(* IEC 61131-3 sources: rusty/tests/lit/multi/external_unit_linkage, 25 files *)

(* ---- interfaces_main.st ---- *)
FUNCTION main : DINT
VAR
    fa : FbA;
    fb : FbB;
END_VAR
    printf('%d$N', call_a(fa));
    printf('%d$N', call_b(fb));
END_FUNCTION

(* ---- properties_c_main.st ---- *)
FUNCTION main : DINT
VAR
    fb : FbExt;
END_VAR
    fb.value := 42;
    printf('%d$N', fb.value);
    printf('%d$N', fb.getValue());
END_FUNCTION

(* ---- properties_main.st ---- *)
FUNCTION main : DINT
VAR
    base : FbBase;
    child : FbChild;
    counter : Counter;
    iface : IValue;
END_VAR
    base.value := 42;
    printf('%d$N', base.value);

    child.value := 5;
    printf('%d$N', child.value);

    printf('%d$N', counter.count);

    iface := child;
    printf('%d$N', iface.value);
END_FUNCTION

(* ---- reference_to_return_lib.st ---- *)
FUNCTION increment : REFERENCE TO DINT
VAR_INPUT
    value : REFERENCE TO DINT;
END_VAR
    value := value + 1;
    increment REF= value;
END_FUNCTION

FUNCTION increment_twice : DINT
VAR
    x : DINT := 5;
    r : REFERENCE TO DINT;
END_VAR
    r REF= x;
    r REF= increment(r);
    r REF= increment(r);
    increment_twice := r;
END_FUNCTION

(* ---- reference_to_return_main.st ---- *)
FUNCTION main : DINT
VAR
    x : DINT := 2;
    r : REFERENCE TO DINT;
END_VAR
    r REF= x;
    r REF= increment(r);
    printf('%d$N', r);
    printf('%d$N', increment_twice());
END_FUNCTION

(* ---- retain_main.st ---- *)
FUNCTION main : DINT
    RetainProgram();
    printf('%d$N', RetainProgram.count);
    printf('%d$N', retainFb.value);
END_FUNCTION

(* ---- retained_fat_pointer_main.st ---- *)
FUNCTION main
    bindA();
    bindB();
    consumerA();
    consumerB();
    printf('%d %d$N', consumerA.result, consumerB.result);
END_FUNCTION

(* ---- retained_fat_pointer_overload_main.st ---- *)
FUNCTION main
    // CHECK: main: done
    printf('main: done$N');
END_FUNCTION

(* ---- retained_fat_pointer_property_main.st ---- *)
FUNCTION main
    VAR
        ownerA : OwnerA;
        ownerB : OwnerB;
    END_VAR
    printf('%d %d$N', ownerA.value, ownerB.value);
END_FUNCTION

(* ---- interface_dispatch_lib.st ---- *)
INTERFACE IShape
    METHOD area : DINT END_METHOD
    PROPERTY_GET name : DINT END_PROPERTY
END_INTERFACE

INTERFACE ISolid EXTENDS IShape
    METHOD volume : DINT END_METHOD
END_INTERFACE

INTERFACE ILogger
    METHOD log : DINT
    VAR_INPUT value : DINT; END_VAR
    END_METHOD
END_INTERFACE

FUNCTION_BLOCK LibSquare IMPLEMENTS IShape
VAR
    side : DINT := 3;
END_VAR
    METHOD area : DINT area := side * side; END_METHOD
    PROPERTY_GET name : DINT name := 100; END_PROPERTY
END_FUNCTION_BLOCK

FUNCTION_BLOCK LibCube EXTENDS LibSquare IMPLEMENTS ISolid
    METHOD volume : DINT volume := area() * side; END_METHOD
    PROPERTY_GET name : DINT name := 200; END_PROPERTY
END_FUNCTION_BLOCK

FUNCTION lib_area_of : DINT
VAR_INPUT shape : IShape; END_VAR
    lib_area_of := shape.area() + shape.name;
END_FUNCTION

FUNCTION_BLOCK LibService
VAR
    logger : ILogger;
    shapes : ARRAY[0..1] OF IShape;
END_VAR
    METHOD inject
    VAR_INPUT l : ILogger; END_VAR
        logger := l;
    END_METHOD

    METHOD add_shape
    VAR_INPUT i : DINT; s : IShape; END_VAR
        shapes[i] := s;
    END_METHOD

    METHOD run : DINT
        run := logger.log(shapes[0].area() + shapes[1].area());
    END_METHOD
END_FUNCTION_BLOCK

FUNCTION lib_volume_as_shape : DINT
VAR_INPUT solid : ISolid; END_VAR
VAR shape : IShape; END_VAR
    shape := solid;
    lib_volume_as_shape := solid.volume() + shape.area();
END_FUNCTION

(* ---- interface_dispatch_main.st ---- *)
FUNCTION_BLOCK AppLogger IMPLEMENTS ILogger
VAR
    last : DINT;
END_VAR
    METHOD log : DINT
    VAR_INPUT value : DINT; END_VAR
        last := value;
        log := value + 1;
    END_METHOD
END_FUNCTION_BLOCK

FUNCTION_BLOCK AppCircle IMPLEMENTS IShape
    METHOD area : DINT area := 7; END_METHOD
    PROPERTY_GET name : DINT name := 300; END_PROPERTY
END_FUNCTION_BLOCK

FUNCTION_BLOCK AppBigCube EXTENDS LibCube
    METHOD area : DINT area := 50; END_METHOD
END_FUNCTION_BLOCK

FUNCTION main : DINT
VAR
    square : LibSquare;
    cube : LibCube;
    bigCube : AppBigCube;
    circle : AppCircle;
    logger : AppLogger;
    service : LibService;
    shape : IShape;
    solid : ISolid;
END_VAR
    // Lib type, called through an interface in the app
    shape := square;
    printf('%d %d$N', shape.area(), shape.name);
    shape := cube;
    printf('%d %d$N', shape.area(), shape.name);
    solid := cube;
    printf('%d$N', solid.volume());

    // App type passed to a lib function that calls through the interface
    printf('%d$N', lib_area_of(circle));
    printf('%d$N', lib_area_of(square));

    // App type that extends a lib type, overriding a method
    shape := bigCube;
    printf('%d %d$N', shape.area(), shape.name);
    printf('%d$N', lib_volume_as_shape(bigCube));

    // Dependency inversion: the lib stores app objects and calls them later
    service.inject(logger);
    service.add_shape(0, circle);
    service.add_shape(1, bigCube);
    printf('%d %d$N', service.run(), logger.last);
END_FUNCTION

(* ---- interfaces_lib_a.st ---- *)
INTERFACE IA
    METHOD a : DINT END_METHOD
END_INTERFACE

FUNCTION_BLOCK FbA IMPLEMENTS IA
    METHOD a : DINT
        a := 1;
    END_METHOD
END_FUNCTION_BLOCK

FUNCTION call_a : DINT
VAR_INPUT
    x : IA;
END_VAR
    call_a := x.a();
END_FUNCTION

(* ---- interfaces_lib_b.st ---- *)
INTERFACE IB
    METHOD b : DINT END_METHOD
END_INTERFACE

FUNCTION_BLOCK FbB IMPLEMENTS IB
    METHOD b : DINT
        b := 2;
    END_METHOD
END_FUNCTION_BLOCK

FUNCTION call_b : DINT
VAR_INPUT
    x : IB;
END_VAR
    call_b := x.b();
END_FUNCTION

(* ---- properties_lib.st ---- *)
INTERFACE IValue
    PROPERTY_GET value : DINT END_PROPERTY
END_INTERFACE

FUNCTION_BLOCK FbBase IMPLEMENTS IValue
VAR
    _value : DINT;
END_VAR
    PROPERTY_GET value : DINT
        value := _value;
    END_PROPERTY

    PROPERTY_SET value : DINT
        _value := value;
    END_PROPERTY
END_FUNCTION_BLOCK

FUNCTION_BLOCK FbChild EXTENDS FbBase
    PROPERTY_GET value : DINT
        value := _value * 2;
    END_PROPERTY
END_FUNCTION_BLOCK

CLASS Counter
VAR
    _count : DINT := 7;
END_VAR
    PROPERTY_GET count : DINT
        count := _count;
    END_PROPERTY
END_CLASS

(* ---- retain_lib.st ---- *)
FUNCTION_BLOCK FbRetain
VAR RETAIN
    value : DINT := 4;
END_VAR
END_FUNCTION_BLOCK

PROGRAM RetainProgram
VAR RETAIN
    count : DINT := 1;
END_VAR
    count := count + 1;
END_PROGRAM

VAR_GLOBAL
    retainFb : FbRetain;
END_VAR

(* ---- retained_fat_pointer_external_app.st ---- *)
INTERFACE IA
    METHOD foo : DINT END_METHOD
END_INTERFACE

{external}
FUNCTION_BLOCK Consumer
VAR_INPUT
    in1 : REFERENCE TO IA;
END_VAR
VAR_OUTPUT
    result : DINT;
END_VAR
END_FUNCTION_BLOCK

{external}
FUNCTION_BLOCK FbA IMPLEMENTS IA
    METHOD foo : DINT END_METHOD
END_FUNCTION_BLOCK

// The declaration keeps the library function's body. Codegen omits it, so the retained fat pointer
// global that the body binds must only be declared here and defined by the library.
{external}
FUNCTION bindExt
VAR_IN_OUT
    consumer : Consumer;
    instance : FbA;
END_VAR
    consumer(instance);
END_FUNCTION

FUNCTION main
VAR
    consumer : Consumer;
    instance : FbA;
END_VAR
    bindExt(consumer, instance);
    consumer();
    printf('%d$N', consumer.result);
END_FUNCTION

(* ---- retained_fat_pointer_external_lib.st ---- *)
INTERFACE IA
    METHOD foo : DINT END_METHOD
END_INTERFACE

FUNCTION_BLOCK Consumer
VAR_INPUT
    in1 : REFERENCE TO IA;
END_VAR
VAR_OUTPUT
    result : DINT;
END_VAR
    result := in1.foo();
END_FUNCTION_BLOCK

FUNCTION_BLOCK FbA IMPLEMENTS IA
    METHOD foo : DINT
        foo := 1;
    END_METHOD
END_FUNCTION_BLOCK

FUNCTION bindExt
VAR_IN_OUT
    consumer : Consumer;
    instance : FbA;
END_VAR
    consumer(instance);
END_FUNCTION

(* ---- retained_fat_pointer_lib_a.st ---- *)
INTERFACE IA
    METHOD foo : DINT END_METHOD
END_INTERFACE

FUNCTION_BLOCK Consumer
VAR_INPUT
    in1 : REFERENCE TO IA;
END_VAR
VAR_OUTPUT
    result : DINT;
END_VAR
    result := in1.foo();
END_FUNCTION_BLOCK

FUNCTION_BLOCK FbA IMPLEMENTS IA
    METHOD foo : DINT
        foo := 1;
    END_METHOD
END_FUNCTION_BLOCK

VAR_GLOBAL
    consumerA : Consumer;
    instanceA : FbA;
END_VAR

FUNCTION bindA
    consumerA(instanceA);
END_FUNCTION

(* ---- retained_fat_pointer_lib_b.st ---- *)
FUNCTION_BLOCK FbB IMPLEMENTS IA
    METHOD foo : DINT
        foo := 2;
    END_METHOD
END_FUNCTION_BLOCK

VAR_GLOBAL
    consumerB : Consumer;
    instanceB : FbB;
END_VAR

FUNCTION bindB
    consumerB(instanceB);
END_FUNCTION

(* ---- retained_fat_pointer_overload_lib_a.st ---- *)
FUNCTION_BLOCK FbOverloadA IMPLEMENTS IA
    METHOD foo : DINT
        foo := 1;
    END_METHOD
END_FUNCTION_BLOCK

VAR_GLOBAL
    overloadConsumerA : Consumer;
    overloadInstanceA : FbOverloadA;
END_VAR

FUNCTION bind<T: ANY_INT> : T
VAR_INPUT
    value : T;
END_VAR
    overloadConsumerA(in1 := overloadInstanceA);
    bind := value;
END_FUNCTION

(* ---- retained_fat_pointer_overload_lib_b.st ---- *)
FUNCTION_BLOCK FbOverloadB IMPLEMENTS IA
    METHOD foo : DINT
        foo := 2;
    END_METHOD
END_FUNCTION_BLOCK

VAR_GLOBAL
    overloadConsumerB : Consumer;
    overloadInstanceB : FbOverloadB;
END_VAR

FUNCTION bind<U: ANY_REAL> : U
VAR_INPUT
    value : U;
END_VAR
    overloadConsumerB(in1 := overloadInstanceB);
    bind := value;
END_FUNCTION

(* ---- retained_fat_pointer_property_lib_a.st ---- *)
FUNCTION_BLOCK FbPropertyA IMPLEMENTS IA
    METHOD foo : DINT
        foo := 1;
    END_METHOD
END_FUNCTION_BLOCK

VAR_GLOBAL
    propertyConsumerA : Consumer;
    propertyInstanceA : FbPropertyA;
END_VAR

FUNCTION_BLOCK OwnerA
    PROPERTY_GET value : DINT
        propertyConsumerA(in1 := propertyInstanceA);
        value := propertyConsumerA.result;
    END_PROPERTY
END_FUNCTION_BLOCK

(* ---- retained_fat_pointer_property_lib_b.st ---- *)
FUNCTION_BLOCK FbPropertyB IMPLEMENTS IA
    METHOD foo : DINT
        foo := 2;
    END_METHOD
END_FUNCTION_BLOCK

VAR_GLOBAL
    propertyConsumerB : Consumer;
    propertyInstanceB : FbPropertyB;
END_VAR

FUNCTION_BLOCK OwnerB
    PROPERTY_GET value : DINT
        propertyConsumerB(in1 := propertyInstanceB);
        value := propertyConsumerB.result;
    END_PROPERTY
END_FUNCTION_BLOCK

(* ---- retained_fat_pointer_template_lib_a.st ---- *)
FUNCTION_BLOCK FbTemplateA IMPLEMENTS IA
    METHOD foo : DINT
        foo := 1;
    END_METHOD
END_FUNCTION_BLOCK

VAR_GLOBAL
    templateConsumerA : Consumer;
    templateInstanceA : FbTemplateA;
END_VAR

FUNCTION bind<T: ANY_INT> : T
VAR_INPUT
    value : T;
END_VAR
    templateConsumerA(in1 := templateInstanceA);
    bind := value;
END_FUNCTION

(* ---- retained_fat_pointer_template_lib_b.st ---- *)
FUNCTION_BLOCK FbTemplateB IMPLEMENTS IA
    METHOD foo : DINT
        foo := 1;
    END_METHOD
END_FUNCTION_BLOCK

VAR_GLOBAL
    templateConsumerB : Consumer;
    templateInstanceB : FbTemplateB;
END_VAR

FUNCTION bind<U: ANY_INT> : U
VAR_INPUT
    value : U;
END_VAR
    templateConsumerB(in1 := templateInstanceB);
    bind := value;
END_FUNCTION
